Fanuc TP program (LS listing): TurnProg.LS

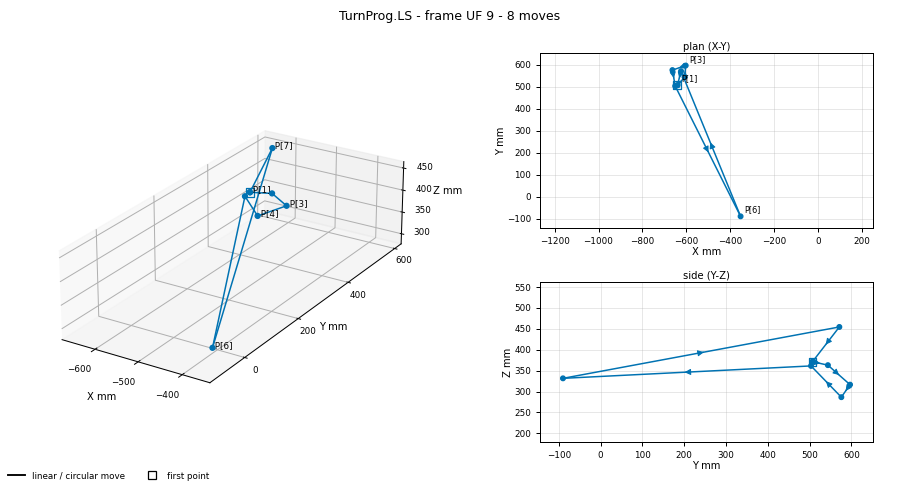
[picture p0: tool path of TurnProg.LS in frame UF 9, 8 of 9 moves have a stored position in this frame; points joined in program order, loops and branches not executed]
/PROG  TurnProg
/ATTR
OWNER		= MNEDITOR;
COMMENT		= "RoboDK sequence";
PROG_SIZE	= 0;
CREATE		= DATE 31-12-14  TIME 12:00:00;
MODIFIED	= DATE 31-12-14  TIME 12:00:00;
FILE_NAME	= TurnProg;
VERSION		= 0;
LINE_COUNT	= 28;
MEMORY_SIZE	= 0;
PROTECT		= READ_WRITE;
TCD:  STACK_SIZE	= 0,
      TASK_PRIORITY	= 50,
      TIME_SLICE	= 0,
      BUSY_LAMP_OFF	= 0,
      ABORT_REQUEST	= 0,
      PAUSE_REQUEST	= 0;
DEFAULT_GROUP	= 1,*,*,*,*,*,*;
CONTROL_CODE	= 00000000 00000000;
/MN
   1:  ! Program generated by RoboDK v6.0.7 for Fanuc ARC Mate 120iD/1 ;
   2:  ! 2L on XX/XX/XXXX 18:00:00 ;
   3:  ! Using nominal kinematics. ;
   4:  PR[9,1]=1234.570 ;
   5:  PR[9,2]=-98.765 ;
   6:  PR[9,3]=50.500 ;
   7:  PR[9,4]=0.000 ;
   8:  PR[9,5]=0.000 ;
   9:  PR[9,6]=30.000 ;
  10:  UFRAME[9]=PR[9] ;
  11:  UFRAME_NUM=9 ;
  12:  PR[9,1]=10.000 ;
  13:  PR[9,2]=20.000 ;
  14:  PR[9,3]=150.000 ;
  15:  PR[9,4]=0.000 ;
  16:  PR[9,5]=0.000 ;
  17:  PR[9,6]=0.000 ;
  18:  UTOOL[9]=PR[9] ;
  19:  UTOOL_NUM=9 ;
  20:L P[1] 200mm/sec FINE ;
  21:L P[2] 200mm/sec FINE ;
  22:L P[3] 200mm/sec FINE ;
  23:L P[4] 200mm/sec FINE ;
  24:L P[5] 200mm/sec FINE ;
  25:L P[6] 200mm/sec FINE ;
  26:L P[7] 200mm/sec FINE ;
  27:L P[8] 200mm/sec FINE ;
  28:J P[9] 20% FINE ;
/POS
P[1]{
   GP1:
    UF : 9, UT : 9,        CONFIG : 'N U T, 1, 0, 0',
	X =  -640.584  mm,	Y =   506.980  mm,	Z =   371.534  mm,
	W =  -165.000 deg,	P =    50.000 deg,	R =   150.000 deg
};
P[2]{
   GP1:
    UF : 9, UT : 9,        CONFIG : 'N U T, 0, -1, 0',
	X =  -607.850  mm,	Y =   543.849  mm,	Z =   363.215  mm,
	W =  -165.000 deg,	P =    50.000 deg,	R =   150.000 deg
};
P[3]{
   GP1:
    UF : 9, UT : 9,        CONFIG : 'F U T, 0, 0, 1',
	X =  -602.951  mm,	Y =   596.788  mm,	Z =   316.595  mm,
	W =  -165.000 deg,	P =    50.000 deg,	R =   150.000 deg
};
P[4]{
   GP1:
    UF : 9, UT : 9,        CONFIG : 'N U B, -1, 0, -1',
	X =  -663.517  mm,	Y =   575.988  mm,	Z =   286.611  mm,
	W =  -165.000 deg,	P =    50.000 deg,	R =   150.000 deg
};
P[5]{
   GP1:
    UF : 9, UT : 9,        CONFIG : 'N D T, 0, 0, 0',
	X =  -650.861  mm,	Y =   503.437  mm,	Z =   361.399  mm,
	W =  -165.000 deg,	P =    50.000 deg,	R =   150.000 deg
};
P[6]{
   GP1:
    UF : 9, UT : 9,        CONFIG : 'F D T, 0, 1, -1',
	X =  -353.026  mm,	Y =   -90.135  mm,	Z =   331.702  mm,
	W =  -169.444 deg,	P =    40.650 deg,	R =   178.023 deg
};
P[7]{
   GP1:
    UF : 9, UT : 9,        CONFIG : 'F D B, 1, -1, 2',
	X =  -624.230  mm,	Y =   571.208  mm,	Z =   454.620  mm,
	W =   -82.711 deg,	P =    44.567 deg,	R =  -122.815 deg
};
P[8]{
   GP1:
    UF : 9, UT : 9,        CONFIG : 'N D B, -1, 1, -2',
	X =  -640.584  mm,	Y =   506.980  mm,	Z =   371.534  mm,
	W =  -165.000 deg,	P =    50.000 deg,	R =   150.000 deg
};
P[9]{
   GP1:
    UF : 9, UT : 9,
	J1=    350.000 deg,	J2=    0.000 deg,	J3=    0.000 deg,
	J4=    -350.000 deg,	J5=    30.000 deg,	J6=    540.000 deg
};
/END
